Fanuc KAREL source: kt00708.KL

-- PROVISIONAL review KL for V1013-1; original PC SHA256 cc49c5c1803e94c7130352aeecf74e3cf9e2c14de2019a66003416b4a7e8c07b
-- Incomplete behavior may be omitted. Consult companion uncertainty JSON. Do not deploy.
PROGRAM KT00708
%NOLOCKGROUP
VAR
  R1 : REAL
  R2 : REAL
  OUT : BOOLEAN
BEGIN
  -- UNRESOLVED_PC offsets 5-16; opcodes 2E,23
  -- UNRESOLVED_PC offsets 21-32; opcodes 2E,23
  -- UNRESOLVED_PC offsets 37-48; opcodes 2E,23
  -- UNRESOLVED_PC offsets 53-64; opcodes 2E,23
  -- UNRESOLVED_PC offsets 69-84; opcodes 22,63,23
  -- UNRESOLVED_PC offsets 89-93; opcodes 7F
END KT00708
